(* IEC 61131-3 sources: JingjiangArm/moonboxpro_arm_8.4/Application/Application/数据类型/系统参数/非保持参数, 3 files *)

(* ---- StGrpParam_UnSave.st ---- *)
(*@CES
Name=StGrpParam_UnSave
Type=Gvl
TypeGuid=2db5746d-d284-4425-9f7f-2663a34b0ebc
Guid=502fdab7-460b-44d8-9c01-902a9f3d20a9
HasDeclaration=True
HasImplementation=False
*)
{DECLARATION}
{attribute 'pack_mode' := '1'}
TYPE StGrpParam_UnSave :
STRUCT
	xCutterOnTop_Uw								: BOOL;(* TRUE=放料上裁 *)
	iDebugVelmpm_AxisA_Uw						: INT;(* A轴调试速度/300m/min *)
	iDebugGirthmm_AxisA_Uw						: INT;(* A轴调试周长/300mm *)
	iDebugVelmpm_AxisB_Uw						: INT;(* B轴调试速度/300m/min *)
	iDebugGirthmm_AxisB_Uw						: INT;(* B轴调试周长/300mm *)
	xCutterOnTop_Rw								: BOOL;(* TRUE=收料上裁 *)
	iDebugVelmpm_AxisA_Rw						: INT;(* A轴调试速度/默认300m/min *)
	iDebugGirthmm_AxisA_Rw						: INT;(* A轴调试周长/默认300mm *)
	iDebugVelmpm_AxisB_Rw						: INT;(* B轴调试速度/默认300m/min *)
	iDebugGirthmm_AxisB_Rw						: INT;(* B轴调试周长/默认300mm *)

	xMachineRev									: BOOL;(* 机器反转 *)

	iPromptMsg									: INT;
	iAlarm_TypeId								: INT;//报警轴的类型
	iAlarm_UnitId								: INT;//报警轴位置
	iIdGSE										: INT;
	xFlag_Stop									: BOOL;(* 停机标志/第1次从当前速度降到空转速度，抬所有色组胶辊/牵引速度到0时抬牵引胶辊，第2次按下则将色组从空转停到0速度 *)
	xFlag_PreStart								: BOOL;(* 预启动标志/从停机状态按(预)启动置位标志 色组速度达到空转速度清xFlag_PreStart标志,置位xFlag_Ink标志;当xFlag_Print标志有效后 *)
	xFlag_Ink									: BOOL;(* 匀墨标志/>20m/min不能联动 *)
	xFlag_InkAccing								: BOOL;(* 匀墨加速中<指0~10m/min那个加速过程> *)
	xFlag_Tension								: BOOL;(* 张力投入标志/张力投入有效时收放料变频开始起作用/收放料就位后按印刷按钮,牵引压辊合压/xFlag_Print有效时张力投入不处理 *)
	xFlag_TensionDone							: BOOL;(* 张力ok，可以投入印刷 *)
	xFlag_Print									: BOOL;(* 张力拉料标志有效时，按联动或印刷按钮 先压收牵(延时2s)再压放牵 印刷标志/印刷色组根据联动标志按用户指定的压辊顺序逐一延时压胶辊/胶辊压合完毕后才可置该标志有效 *)
	xFlag_Estop									: BOOL;(* 急停标志/和停机一样要减速到0，只不过减速时间是急停时间 *)
	xFlag_AutoAcc								: BOOL;(* 自动加速 *)
	xFlag_AutoDec								: BOOL;(* 自动减速 *)
	xFlag_ManuAcc								: BOOL;(* 手动加速 *)
	xFlag_ManuDec								: BOOL;(* 手动减速 *)
	xFlag_Accing								: BOOL;(* 加速中 *)
	xFlag_Decing								: BOOL;(* 减速中 *)
	xFlag_EStoping								: BOOL;(* 正在急停中 *)
	xFlag_Stoping								: BOOL;(* 停机中 *)
	xFlag_GotoInking							: BOOL;(* 转到匀墨 *)
	xFlag_InPressing							: BOOL;(* 顺序压辊中 *)
	xFlag_RollerPressDone						: BOOL;(* 压辊处理完成 *)
	xFlag_InchRun								: BOOL;(* 至少有1色处于单运行 *)
	xFlag_AllInchRun							: BOOL;(* 整机单运行标志 *)
	xFlag_AllPress								: BOOL;(* 全体合压 *)
	xFlag_AllUnpress							: BOOL;(* 全体离压 *)
	xFlag_RollerPressAtLeast1					: BOOL;(* 至少1色色组合压 *)
	axFlag_PrnLen_Alarm							: ARRAY [1..3] OF BOOL;(* 计长报警标志 *)
	xFlag_LinkageAxisAlarm						: BOOL;(* 至少有1个联动轴发生报警 *)
	xFlag_TensionUnfinished						: BOOL;(* 张力未完成 *)
	xFlag_VelTooHigh							: BOOL;(* 速度过高 *)
	xFlag_PrestartTimeout						: BOOL;(* 预启动超时标志 *)
	xFlag_KeepAlarming							: BOOL;(* 维持报警*)
	xFlag_ArrivedToTargetVel					: BOOL;(* 到达目标速度 *)
	xFlag_FilmAccDecDone						: BOOL;(* 料膜加减速完成 *)
	xSlowStopTenEn								: BOOL;(* 收放料慢速松料使能/TRUE *)
	xIsDebugMode_Machine						: BOOL;(* 机器调试模式 *)
	uiFilmThickNess								: UINT;(* 料膜厚度/20微米 *)
	abyClrPrnLenCount_Rw						: ARRAY [1..3] OF BYTE;

	iTimeSec_AccDec_AllTheWay					: INT;(* 全程加减速所需要的秒 *)
	rAccDecTime_ThisTime						: REAL;(* 本次加减速时间/单位:s *)

(*2021.11.5.084313/								/ 用于界面显示标准卷径信息 *)
	alrStdVol_Diam_Axis_Hmi						: ARRAY [1..4] OF LREAL;(* 标准卷径值| *)
	alrStdVol_Volt_Axis_Hmi						: ARRAY [1..4] OF LREAL;(* 标准卷径对应的电压值|2019.1.25.142552|更名A轴 *)
	alrStdVol_Coef_Axis_Hmi						: ARRAY [0..4] OF LREAL;(* 分段系数|2019.1.25.142601|更名A轴|[0]表<=1,[1]表>1&& <=2,[2]表>2&& <=3,[3]表>3&& <=4,[4]表>4 *)

	(* 速度 *)
	rVel_Cur									: REAL;(* 当前速度/单位:m/min *)
	rVel_Cur_HMI								: REAL;
	rVel_Film									: REAL;(* 料膜速度/0 *)
	(*											/放料部分 *)
	iSid_AxisA_Uw								: INT;(* 放料站id/-1表示变频/2021.11.21.192354/hdp *)
	xStationOnline_AxisA_Uw						: BOOL;(* 放料a轴驱动器在线标志/2021.12.4.175524/hdp *)
	xMotRev_AxisA_Uw							: BOOL;(* TRUE.放料运动反向/2021.11.21.192354/hdp *)

	iSid_AxisB_Uw								: INT;(* 放料站id/-1表示变频/2021.11.21.192354/hdp *)
	xStationOnline_AxisB_Uw						: BOOL;(* 放料b轴驱动器在线标志/2021.12.4.175524/hdp *)
	xMotRev_AxisB_Uw							: BOOL;(* TRUE.放料运动反向/2021.11.21.192354/hdp *)

	rAI_Uw										: REAL;(* 放料摆臂模拟量输入/-中位值 *)
	rAI_Act_Uw									: REAL;(* 放料摆臂实际模拟量值/2021.11.18.210606 *)
	rAI_HMI_Uw									: REAL;(* 放料摆臂值显示用 *)
	rAI_DiamMeasure_Uw							: REAL;(* 放料卷径测量输入反馈 *)
	arKpid_Current_Uw							: ARRAY [1..3] OF REAL;(* 当前放料pid监控 *)
	stStTimeSet_DnCut_UpCut_Uw_Hmi				: StTimeSet_DnCut_UpCut;(* 放料端的裁切时间集/界面显示 *)
	arKpid_Current_Rw							: ARRAY [1..3] OF REAL;(* 当前收料pid监控 *)
	stStTimeSet_DnCut_UpCut_Rw_Hmi				: StTimeSet_DnCut_UpCut;(* 收料端的裁切时间集/界面显示 *)
	rVel_PreDrv_Uw								: REAL;(* 放料预驱速度 *)
	xReflectionSensorValid_Uw					: BOOL;(* 放料使用弧面信号/FALSE *)
	xReflectSensorLoss_Uw						: BOOL;(* 放料弧面信号丢失标志/FALSE *)
	rDiam_NewVol_Uw								: REAL;(* 放料新卷卷径 *)
	rTowerThetaCur_Uw							: REAL;(* 翻转架当前弧度/0 *)
	rFilmToTowerRollerDis_Uw				: REAL;(*料膜距离导向辊距离|mm*)
	xFilmTouchRoller_Uw						: BOOL;(*料膜接触到了辊子标志*)

	xSts_PreCutting_Uw							: BOOL;(* 放料预备接料/FALSE *)
	rDebugCurVelmpmAxisA_Uw						: REAL;(* A轴调试当前速度/m/min *)
	rDebugCurVelrpmAxisA_Uw						: REAL;(* A轴调试当前速度/r/min *)
	rDebugCurVelmpmAxisB_Uw						: REAL;(* B轴调试当前速度/m/min *)
	rDebugCurVelrpmAxisB_Uw						: REAL;(* B轴调试当前速度/r/min *)

	rDeltaW_RPMIN_Uw							: REAL;(* 放料翻转架转动时候的转速补偿值/0 *)
	xDebugMode_AbsEnc_Uw						: BOOL;(* 放料绝对值编码器调试模式/FALSE *)
	dwAbsEncSinglePos_Uw						: DWORD;(* 放料单圈位置/0 *)
	dwAbsEncSPos_Cur_Uw							: DWORD;(* 放料当前绝对位置/0 *)

	byEncodeValueWr_Uw							: BYTE;(* 放料编码器值写入/放料:01写入轴定位值/02写入A轴最小径定位值/0 *)
	rAIByAbsEnc_Cur_Uw							: REAL;(* 放料绝对值编码器位置转换的电压值/0 *)
	xCutterOnTopFroDebug_Uw						: BOOL;(* 放料上裁刀标志/用于调试/FALSE *)
	xCurAxisAFroDebug_Uw						: BOOL;(* 放料预驱轴为A轴标志/用于调试/FALSE *)
	xAlarmBell_Uw								: BOOL;(* 放料响铃常输出/用于控制定位写入响铃提示使用/FALSE *)
	xIsDebug_DiaMeasure_Uw						: BOOL;(* 放料卷径测量调试模式标志/FALSE *)
	byIsDebug_DiaMeasureArea_Uw					: BYTE;(* 放料卷径测量调试的时候卷径区域值/1 *)
	xIsDebuging_DiaMeasure_Uw					: BOOL;(* 放料卷径测量调试中/FALSE *)
	xCancelDebuging_DiaMeasure_Uw				: BOOL;(* 放料取消卷径测量调试中/FALSE *)
	byAxisDebugBit_Uw							: BYTE;(* 放料轴调试标志/.0\调试使能.1\A轴调试运行.2\A轴自动加减速.3\A轴运行中.4\B轴调试运行.5\B轴自动加减速.6\B轴运行中/0 *)
	byAxisDebugBit_Uw_2							: BYTE;(* 放料2轴调试标志/.0\调试使能.1\A轴调试运行.2\A轴自动加减速.3\A轴运行中.4\B轴调试运行.5\B轴自动加减速.6\B轴运行中/0 *)
	xEnCodeErr_Uw								: BOOL;(* 放料编码器故障*)
	xEnCodeErr_Rw								: BOOL;(* 收料编码器故障*)

	rPi_Value_Uw								: REAL;(* 放料pi值/0 *)
	rForwardStep_Uw								: REAL;(* 放料升降速前馈/0 *)
	rTotalPiValue_Uw							: REAL;
	xAxisAForeward_Uw							: BOOL;(* 放料A轴正转/FALSE *)
	xAxisBForeward_Uw							: BOOL;(* 放料B轴正转/FALSE *)
	rVelRPM_Cur_Uw								: REAL;(* 放料当前转速/0 *)
	rAxisAVelRPM_Cur_Uw							: REAL;(* 放料A轴转速/0/2021.11.18.201209 *)
	rAxisBVelRPM_Cur_Uw							: REAL;(* 放料B轴转速/0/2021.11.18.201209 *)
	xFlag_DiamCalc_ing_Uw						: BOOL;(* 放料卷径计算中 *)
	xFlag_DiamCalc_end_Uw						: BOOL;(* 放料卷径计算完成 *)
	xFlag_DiamMeasure_end_Uw					: BOOL;(* 放料卷径测量完成 *)
	xFlag_PreDrv_ing_Uw							: BOOL;(* 放料预驱中... *)
	xFlag_PreDrv_end_Uw							: BOOL;(* 放料预驱完成  *)
	xFlag_Cut_ing_Uw							: BOOL;
	xFlag_Cut_end_Uw							: BOOL;
	xFlag_VolDiamAlarm_Uw						: BOOL;(* 卷径报警标志 *)
	rAI_DiamMeasure_HMI_Uw						: REAL;(* 兼容摆臂输入类型转换后的卷径测量结果屏显值/2021.11.5.175329 *)
	xAITypeBtn_Uw								: BOOL;(* 输入类型切换按钮/2021.11.18.201254 *)

	(*											/收料部分 *)
	iSid_AxisA_Rw								: INT;(* 收料站id/-1表示变频/2021.11.21.192354/hdp *)
	xStationOnline_AxisA_Rw						: BOOL;(* 收料a轴驱动器在线标志/2021.12.4.175524/hdp *)
	xMotRev_AxisA_Rw							: BOOL;(* TRUE.收料运动反向/2021.11.21.192354/hdp *)

	iSid_AxisB_Rw								: INT;(* 收料站id/-1表示变频/2021.11.21.192354/hdp *)
	xStationOnline_AxisB_Rw						: BOOL;(* 收料b轴驱动器在线标志/2021.12.4.175524/hdp *)
	xMotRev_AxisB_Rw							: BOOL;(* TRUE.收料运动反向/2021.11.21.192354/hdp *)

	rAI_Rw										: REAL;(* 收料摆臂模拟量输入/-中位值 *)
	rAI_Act_Rw									: REAL;(* 收料摆臂实际模拟量值/2021.11.18.201450 *)
	rAI_HMI_Rw									: REAL;(* 收料摆臂值显示用 *)
	rVel_PreDrv_Rw								: REAL;(* 收料预驱速度 *)
	rDiam_NewVol_Rw								: REAL;(* 收料新卷卷径 *)
	rTaper_Rw									: REAL;(* 收料锥度 *)

	xSts_PreCutting_Rw							: BOOL;(* 收料预备接料 *)
	rDebugCurVelmpmAxisA_Rw						: REAL;(* A轴调试当前速度/m/min *)
	rDebugCurVelrpmAxisA_Rw						: REAL;(* A轴调试当前速度/r/min *)

	rDebugCurVelmpmAxisB_Rw						: REAL;(* B轴调试当前速度/m/min *)
	rDebugCurVelrpmAxisB_Rw						: REAL;(* B轴调试当前速度/r/min *)
	xDebugMode_AbsEnc_Rw						: BOOL;(* 收料绝对值编码器调试模式/默认FALSE *)
	dwAbsEncSinglePos_Rw						: DWORD;(* 收料单圈位置/0 *)
	dwAbsEncSPos_Cur_Rw							: DWORD;(* 收料当前绝对位置/0 *)
	byEncodeValueWr_Rw							: BYTE;(* 收料编码器值写入/收料/01写入轴定位值/0 *)
	xCutterOnTopFroDebug_Rw						: BOOL;(* 收料上裁刀标志/用于调试/FALSE *)
	xCurAxisAFroDebug_Rw						: BOOL;(* 收料预驱轴为A轴标志/用于调试/FALSE *)
	x6InchFroDebug_Rw       					: BOOL;(* 收料6寸标志/用于调试/FALSE*)
	xAlarmBell_Rw								: BOOL;(* 收料响铃常输出/用于控制定位写入响铃提示使用/FALSE *)
	byAxisDebugBit_Rw							: BYTE;(* 收料轴调试标志/.0\调试使能.1\A轴调试运行.2\A轴自动加减速.3\A轴运行中.4\B轴调试运行.5\B轴自动加减速.6\B轴运行中/0 *)
	rPi_Value_Rw								: REAL;(* 收料pi值/0 *)
	rForwardStep_Rw								: REAL;(* 收料升降速前馈/0 *)
	rTotalPiValue_Rw							: REAL;
	xAxisAForeward_Rw							: BOOL;(* 收料A轴正转/FALSE *)
	xAxisBForeward_Rw							: BOOL;(* 收料B轴正转/FALSE *)
	rVelRPM_Cur_Rw								: REAL;(* 收料当前转速/0 *)
	rAxisAVelRPM_Cur_Rw							: REAL;(* 收料A轴转速/0/2021.11.18.201604 *)
	rAxisBVelRPM_Cur_Rw							: REAL;(* 收料B轴转速/0/2021.11.18.201608 *)
	xFlag_6Inch_Rw								: BOOL;(* 收料6寸标志/反之为3寸/FALSE *)
	xFlag_PreDrv_ing_Rw							: BOOL;(* 收料预驱中... *)
	xFlag_PreDrv_end_Rw							: BOOL;(* 收料预驱完成 *)
	xFlag_Cut_ing_Rw							: BOOL;(* 收料裁切中 *)
	xFlag_Cut_end_Rw							: BOOL;(* 收料裁切完成 *)
	xAITypeBtn_Rw								: BOOL;(* 输入类型切换按钮 *)

	(*											/放牵部分 *)
	iSid_If										: INT;(* 放牵站id/-1表示变频 *)
	xStationOnline_If							: BOOL;(* 放牵驱动器在线标志/2021.12.4.175524/hdp *)
	xMotRev_If									: BOOL;(* TRUE.放牵运动反向/2021.11.16.134652/+ *)
(* 2021.12.29.153030/hdp *)

	rAI_If										: REAL;(* 放牵摆臂模拟量输入/-中位值 *)
	rAI_Act_If									: REAL;(* 放牵摆臂实际模拟量值/2021.11.18.201802 *)
	rAI_HMI_If									: REAL;(* 放牵摆臂值显示用 *)
	xInchBtn_If									: BOOL;(* 放牵单运行/FALSE *)
	xRollerSts_If								: BOOL;(* 放牵压辊/FALSE *)
	xRunEn_If									: BOOL;(* 放牵运动使能/0/2021.11.18.201925 *)
	rVel_Cur_If									: REAL;(* 放牵速度/0 *)
	rPi_Value_If								: REAL;(* 放牵pi值/0 *)
	rForwardStep_If								: REAL;(* 放牵升降速前馈/0 *)
	rUsingGirth_If								: REAL;(* 放牵速度控制实际使用的周长/500mm *)
	xInching_If									: BOOL;(* 放牵单运行中/FALSE *)
	xAITypeBtn_if								: BOOL;(* 输入类型切换按钮 *)
	(*											/收牵部分 *)
	iSid_Of										: INT;(* 收牵站id/-1表示变频 *)
	xStationOnline_Of							: BOOL;(* 收牵驱动器在线标志/2021.12.4.175524/hdp *)
	xMotRev_Of									: BOOL;(* TRUE.收牵运动反向/2021.11.16.134652/+ *)

	rAI_Of										: REAL;(* 收牵摆臂模拟量输入/-中位值 *)
	rAI_Act_Of									: REAL;(* 收牵摆臂实际模拟量值/2021.11.18.202051 *)
	rAI_HMI_Of									: REAL;(* 收牵摆臂值显示用 *)
	xInchBtn_Of									: BOOL;(* 收牵单运行/FALSE *)
	xRollerSts_Of								: BOOL;(* 收牵压辊/FALSE *)
	xRunEn_Of									: BOOL;(* 收牵运动使能/0/2021.11.18.202215 *)
	rVel_Cur_Of									: REAL;(* 收牵速度/0 *)
	rPi_Value_Of								: REAL;(* 收牵pi值/0 *)
	rForwardStep_Of								: REAL;(* 收牵升降速前馈/0 *)
	rUsingGirth_Of								: REAL;(* 收牵速度控制实际使用的周长/500mm *)
	xInching_Of									: BOOL;(* 收牵单运行中/FALSE *)
	xAITypeBtn_Of								: BOOL;(* 输入类型切换按钮/2021.11.18.202322 *)
	sCurRecipeName_InUse							: STRING ;(*当前加在的配方*)
	dwSTS_ALL									: DWORD;(* 2021.11.4.174929 *)
(*												/ 整机状态 *)
(*												/bit0.整机套印纵向自动 *)
(*												/bit1.整机套印横向自动 *)
(*												/*)
(*												/bit8.主站的通讯记录到日志中 *)
(*												/*)
(*												/*)
(*												/bit16.主站请置该标志有效/2021.11.6.102700 *)
(*												/bit17.置位标识显示精采样波形 *)
(*												/*)
(*												/*)
(*												/*)
(*												/bit24.dll显示调试信息/2021.12.1.191835/hdp *)
(*												/bit25.精采样显示阀值3 *)
(*												/bit26.精采样显示阀值2 *)
(*												/bit27.精采样显示阀值1 *)
(*												/bit28.精采样显示峰值位置 *)
(*												/bit29.精采样显示最小值位置 *)
(*												/bit30.精采样显示最大值位置 *)
(*												/bit31.精采样显示基线 *)

	xAutoAccDec_Hmi								: BOOL;
	xFlag_IfOf_Ink								: BOOL;(*空转牵引联动标志*)
	xFlag_FastStoping						: BOOL;
	rFinalVelocity							: REAL;(*末速度*)

	xFlag_AutoMaticCutting_Uw					: BOOL;(*2022.4.25.090246 自动裁切中标志*)
(*	abyReserved1							: ARRAY [1..4] OF BYTE;*)
	xFlag_AutoMaticCutting_rw					: BOOL;(*2022.4.25.090246 自动裁切中标志*)
	rAutoMaticCuttingLenth_CurMode_uw			: REAL;(*放料自动裁切当前模式下的计米值|2022.4.26.101850*)
	rActRemainFilmLenth_Uw						: REAL;(*实际剩余长度|mm-测量值*)
	rAutoMaticCuttingLenth_CurMode_Rw			: REAL;(*收料自动裁切当前模式下的计米值|2022.4.26.101850*)

	xCurAxisDia_Uw_Wr							: BOOL;(*写入当前轴的卷径|2022.4.9.230449*)
	xCurAxisDia_Rw_Wr							: BOOL;(*写入当前轴的卷径|2022.4.9.230449*)
	rTaper_Cur_Uw								: REAL;(*锥度当前|放料|*)
	rTaper_Cur_If								: REAL;(*锥度当前|放牵|*)
	rTaper_Cur_Of								: REAL;(*锥度当前|收牵|*)

	rTaperValueBegin_Hmi_Uw						: REAL;(*放料起始锥度显示值|根据单位切换*)
	rTaperValueEnd_Hmi_Uw						: REAL;(*放料结束锥度显示值|根据单位切换*)
	rTaperValueBegin_Hmi_Rw						: REAL;(*收料起始锥度显示值|根据单位切换*)
	rTaperValueEnd_Hmi_Rw						: REAL;(*收料结束锥度显示值|根据单位切换*)
	rTaperValueBegin_Hmi_If						: REAL;(*放牵起始锥度显示值|根据单位切换*)
	rTaperValueEnd_Hmi_If						: REAL;(*放牵结束锥度显示值|根据单位切换*)
	rTaperValueBegin_Hmi_Of						: REAL;(*收牵起始锥度显示值|根据单位切换*)
	rTaperValueEnd_Hmi_Of						: REAL;(*收牵结束锥度显示值|根据单位切换*)

	byTaperUnitConfirm_Uw						: BYTE;(*放料锥度单位确认|.0 N确认|.1 Mpa确认*)
	byTaperUnitConfirm_Rw						: BYTE;(*收料锥度单位确认|.0 N确认|.1 Mpa确认*)
	byTaperUnitConfirm_If						: BYTE;(*放牵锥度单位确认|.0 N确认|.1 Mpa确认*)
	byTaperUnitConfirm_Of						: BYTE;(*收牵锥度单位确认|.0 N确认|.1 Mpa确认*)
	(*2021.7.29.105859 增加|16BYTES*)
	rTaperValueCur_Hmi_If						: REAL;(*放牵锥度当前值|根据单位切换*)
	rTaperValueCur_Hmi_of						: REAL;(*收牵锥度当前值|根据单位切换*)
	rTaperValueCur_Hmi_Uw						: REAL;(*放料锥度当前值|根据单位切换*)
	rTaperValueCur_Hmi_Rw						: REAL;(*收料锥度当前值|根据单位切换*)
	rValue_DiaMeasure							: REAL;(*卷径测量采样值*)
	rVolt_CalcDiam_Used_Watch					: REAL;(*计算卷径的电压值*)
	rAO_Inverter_Uw_AxisA						: REAL;(*放料A轴输出|2017-08-12 17:25:33*)
	rAO_Inverter_Uw_AxisB						: REAL;(*放料B轴输出|2017-08-12 17:25:33*)
	rAO_Inverter_Rw_AxisA						: REAL;(*收料A轴输出|2017-08-12 17:25:33*)
	rAO_Inverter_Rw_AxisB						: REAL;(*收料B轴输出|2017-08-12 17:25:33*)

	xBtn_HorzPreRegister_Repeat				: BOOL;(*横向重复值按钮*)
	xBtn_HorzPreRegister_Setup				: BOOL;(*横向设定值按钮*)
	xSts_HorzPreRegister					: BOOL;(*横向预套准状态*)
	xMode_HorzPreRegister					: BOOL;(*横向预套准方式：FALSE为设定值;TRUE是重复值*)
	xFlag_HorzPreRegister_All_end			: BOOL;(*横向预套准全部完成*)
	xFlag_Home								: BOOL;
	xFlag_Home_ing							: BOOL;
	xFlag_Home_end							: BOOL;
	xFlag_ConfirmPreRegHomePos				: BOOL;(*2017-09-13 12:51:52| 确认预套准基准点*)
	xFlag_ConfirmPreRegHomePos_ing			: BOOL;(*确认预套准基准点-ing*)
	xFlag_ConfirmPreRegHomePos_end			: BOOL;(*确认预套准基准点-end*)
	xFlag_PreRegister						: BOOL;
	xFlag_PreRegister_ing					: BOOL;
	xFlag_PreRegister_end					: BOOL;
	xFlag_PhaseRestore						: BOOL;(*相位恢复*)
	xFlag_PhaseRestore_ing					: BOOL;(*相位恢复-ing*)
	xFlag_PhaseRestore_end					: BOOL;(*相位恢复-end*)
	xBtn_Home								: BOOL;
	xBtn_ConfirmPreRegHomePos				: BOOL;
	xBtn_PreRegister						: BOOL;
	xBtn_PhaseSave							: BOOL;(*相位保存*)
	xBtn_PhaseRestore						: BOOL;(*相位恢复*)
	xFlag_MotionParamInitialized				: BOOL;(*加速度初始化完成-计算加速度目标速度加加速度*)
	xFlag_AccDecStop							: BOOL;
	//下面时牵引收放料中心辊的离线报警位置偏差报警标志
	xNetOffline_CENTRAL:BOOL;
	xAxisAlarm_CENTRAL:BOOL;
	xPosDeviationAlarm_CENTRAL:BOOL;
	xNetOffline_CENTRAL2:BOOL;
	xAxisAlarm_CENTRAL2:BOOL;
	xPosDeviationAlarm_CENTRAL2:BOOL;
	xNetOffline_IF:BOOL;
	xAxisAlarm_IF:BOOL;
	xPosDeviationAlarm_IF:BOOL;
	xNetOffline_OF:BOOL;
	xAxisAlarm_OF:BOOL;
	xPosDeviationAlarm_OF:BOOL;
	xNetOffline_UW_A:BOOL;
	xAxisAlarm_UW_A:BOOL;
	xPosDeviationAlarm_UW_A:BOOL;
	xNetOffline_UW_B:BOOL;
	xAxisAlarm_UW_B:BOOL;
	xPosDeviationAlarm_UW_B:BOOL;
	xNetOffline_RW_A:BOOL;
	xAxisAlarm_RW_A:BOOL;
	xPosDeviationAlarm_RW_A:BOOL;
	xNetOffline_RW_B:BOOL;
	xAxisAlarm_RW_B:BOOL;
	xPosDeviationAlarm_RW_B:BOOL;
	//2023.8.18.143718具体报警信息
	dwAlarmDetail_CENTRAL:DWORD;//轴报警信息-ZHONGX
	dwAlarmDetail_CENTRAL2:DWORD;//轴报警信息-ZHONGX

	dwAlarmDetail_IF:DWORD;//轴报警信息-放牵
	dwAlarmDetail_OF:DWORD;//轴报警信息-收前
	dwAlarmDetail_UW_A:DWORD;//轴报警信息-放A
	dwAlarmDetail_UW_B:DWORD;//轴报警信息-放B
	dwAlarmDetail_RW_A:DWORD;//轴报警信息-收A
	dwAlarmDetail_RW_B:DWORD;//轴报警信息-收B

	xValid_CentralDrum							: BOOL;(* 中心滚筒有效标志 *)
	iSid_CentralDrum							: INT;(* 中心滚筒站id/初始-1/有效性通过查表确定 *)
	xStationOnline_CentralDrum					: BOOL;(* 站在线标志-中心滚筒/读取站号以后实时更新 *)
	xMotRev_CentralDrum							: BOOL;(* 中心滚筒电机反向运动 *)
	rAxisVel_CentralDrum						: REAL;(* 中心滚筒轴速度 *)
	xPrintInching: BOOL;//整机点动
	rVel_Inching_Print: REAL;//点动速度
	xTapPosition_Breaking					: BOOL;(*断料档位|*)
	xTapPosition_UniformInk					: BOOL;(*匀墨档位|*)
	xTapPosition_Printing					: BOOL;(*印刷档位|*)
	wEn_UwRw_IfOf_Center					: WORD;(*牵引收放料中心辊的使能标志*)
											(*bit0:放牵*)
											(*bit1:收牵*)
											(*bit2:放A*)
											(*bit3:放B*)
											(*bit4:收A*)
											(*bit5:收B*)
											(*bit6:中心辊1*)
											(*bit7:中心辊2*)
	aiMotionStep_AllStation					: ARRAY [1..MAX_STATION_NUM] OF INT;
	byBtn_ConfirmMedian						: BYTE;
	xUwVolDiamMeasurementFailed								: BIT;(*放料卷径检测失败*)
	xBtnClrAlarmInf											: BIT;(*报警清楚按钮*)

	byPseudoRandomId						: BYTE:=1;(*=0 放牵|=1 放料|=2 收料 |=3 收牵*)
	xPseudoRandomEn							: BOOL;(*伪随机使能*)
	aiTestPseudoRandom_Kp					: ARRAY [1..3] OF INT;(*伪随机测试Kp*)
	aiTestPseudoRandom_Kd					: ARRAY [1..3] OF INT;(*伪随机测试Kd*)
	xPseudoRandomTsting						: BOOL;(*伪随机测试中*)
	xDebug_Enc_Uw							: BOOL;(*放料调试*)
	xDebug_Enc_Rw							: BOOL;(*收料调试*)
	wAxisDebug_UwRw							: WORD;(*轴调试标志|.0\放料调试使能.1\放料A轴调试运行.2\放料A轴自动加减速.3\放料A轴运行中.4\放料B轴调试运行.5\放料B轴自动加减速.6\放料B轴运行中
									  .8\收料调试使能.9\收料A轴调试运行.10\收料A轴自动加减速.11\收料A轴运行中.12\收料B轴调试运行.13\收料B轴自动加减速.14\收料B轴运行中*)
	xFlag_SafeTyGratingProctec_Uw			: BOOL;(*放料光栅保护标志*)
	xFlag_SafeTyGratingProctec_Rw			: BOOL;(*放料光栅保护标志*)

	bySetTestPid_IfOf:BYTE;(*设置伪随机测试的pid值*)
	bySetTestPid_Uw:BYTE;(*设置伪随机测试的pid值*)
	bySetTestPid_Rw:BYTE;(*设置伪随机测试的pid值*)
	bySetTestPid_If:BYTE;(*设置伪随机测试的pid值*)
	bySetTestPid_Of:BYTE;(*设置伪随机测试的pid值*)
	xLinkage_IfOf_Ink: BOOL;
	xFlag_Cut_end_Uw_UseInOtherPrg: BOOL;
	xFlag_Cut_ing_Uw_UseInOtherPrg: BOOL;
	xFlag_Cut_end_Rw_UseInOtherPrg: BOOL;
	xConfirmRad0: BOOL;(*0弧度确认*)
	xFlag_Follow_1U_V_UwCut		: BOOL;(*裁切跟一色标志*)
	xKeepAlarm_NoMaterial			: BOOL;(*没料持续报警*)
	xKnob_6Inch_Rw				: BOOL;(*界面收料6吋切换开关*)
	xWillAutoMaticPreCut_Uw		: BOOL;(**)
	axMeasure_StdVol						: ARRAY [1..4] OF BOOL;(*卷径测量按钮*)
	rPseudoRandomRoundAmplitude_Cur		: REAL;

	rAxisAFreq_Uw						: REAL;(*放料A频率监控*)
	rAxisBFreq_Uw						: REAL;(*放料A频率监控*)
	rAxisAFreq_Rw						: REAL;(*放料A频率监控*)
	rAxisBFreq_Rw						: REAL;(*放料A频率监控*)

	xAllowSwitchCutter_Uw				: BOOL;(*收放料允许切换上下裁刀标志@|./0 放料可以|./1 收料可以*)
	xAllowSwitchCutter_Rw				: BOOL;(*收放料允许切换上下裁刀标志@|./0 放料可以|./1 收料可以*)
	xAxisALocation_Use_Uw					: BOOL;
	xAxisBLocation_Use_Uw					: BOOL;
	xAxisALocation_Use_Rw					: BOOL;
	xAxisBLocation_Use_Rw					: BOOL;

	rWuCompensate_Uw:REAL;(*补偿的转速(R/MIN)|计算的*)
	rWuCompensate_Act_Uw:REAL;(*补偿的转速(R/MIN)|实际使用的*)

	rWuCompensate_Rw:REAL;(*补偿的转速(R/MIN)|计算的*)
	rWuCompensate_Act_Rw:REAL;(*补偿的转速(R/MIN)|实际使用的*)
	rTaperMax_Uw: REAL;
	rTaperMax_Rw: REAL;
	rTaperMax_If: REAL;
	rTaperMax_Of: REAL;

	xGirthCalFinish_If: BOOL;
	xGirthCalFinish_Of: BOOL;
	(*扰动输出的控制输入参数@2024.12.3.102359*)
	xEn_Disturbance_If: BOOL;(*扰动使能*)
	rFreq_Disturbance_If: REAL:=1;(*扰动频率@hz*)
	rAmplitude_Disturbance_If:REAL:=1;(*扰动幅值*)
	uiTotalTime_Disturbance_If: UINT:=0;(*扰动输出的总时间|=0 代表一直输出@s*)
	xOuting_sin_If:BOOL:=FALSE;(*输出标志*)
	rResult_sin_If: REAL:=0;
	xEn_Disturbance_Of: BOOL;(*扰动使能*)
	rFreq_Disturbance_Of: REAL:=1;(*扰动频率@hz*)
	rAmplitude_Disturbance_Of:REAL:=1;(*扰动幅值*)
	uiTotalTime_Disturbance_Of: UINT:=0;(*扰动输出的总时间|=0 代表一直输出@s*)
	xOuting_sin_Of:BOOL:=FALSE;(*输出标志*)
	rResult_sin_Of: REAL:=0;
	rVelRPM_Cur_If: REAL;(*放牵转速*)
	rVelRPM_Cur_Of: REAL;(*收牵转速*)
	byPseudoRandomRoundTimes_Cur: BYTE;(*伪随机测试当前次数*)
	xFlagFollow1U_AccDecing: BOOL;(*加减速跟踪第一色标志*)
	byGrpArcAxisNum			: BYTE;
	abyGrpArcAxisList: ARRAY [1..MAX_UNIT_NUM] OF BYTE;
	abyGrpFollowArcIdList: ARRAY [1..MAX_UNIT_NUM] OF BYTE;
	abyGrpArcIdList	: ARRAY [1..MAX_UNIT_NUM] OF INT;
	xEnaTestARC_Ink							: BOOL;(*空转测试使能*)
	rAcceleration_Max				: REAL;(*最大加速度*)
	rAcceleration_Cur				: REAL;(*当前加速度*)

	byGrpAxisNum_Pu					: BYTE;
	abyGrpAxisList					: ARRAY [1..MAX_UNIT_NUM] OF BYTE;
	iAxisId_StepTest_V						: INT;(*阶跃测试的轴id*)
	iMicron_StepTest1_V						: INT;(*阶跃测试的数值|单位:um*)
	iMicron_StepTest2_V						: INT;(*阶跃测试的数值|单位:um*)
	iInterval_StepTest12					: INT;(*2此阶跃的间隔|幅*)

	xSwitch_AutoAdjust_V_Grp				: BIT;(*整机手自动*)
	xSwitch_AutoAdjust_H_Grp				: BIT;(*整机手自动*)
	xLinkage_If								: BIT;(*放牵联动*)
	xLinkage_Of								: BIT;(*收牵联动*)
	xMoveEnable_Motor_If					: BIT;
	xMoveEnable_Motor_Of					: BIT;
	rMainVel_Uw : REAL;
	rMainVel_Rw : REAL;

	(*2025.8.13.103441||新增工艺参数*)
	lrAxisScraperVel:LREAL;
	rHz_UnitScraper_CurrWR: REAL;(*刮刀速度写入变频值-485变频*)
	rHz_UnitInkRoller_CurrWR: REAL;

	(*2025.08.13.145324 || 至少联动一色标志*)
	xFlag_LinkageAtleast1Axis					: BOOL;
	(*新增变量-开始|wang.nt|2025.08.13.144038*)
	xWillAutoMaticPreCut_Rw : BOOL;(*收料即将自动接料*)
	xFlag_HotBlowerStopDelay : BOOL;(*热风延时关闭中*)
	xInverterAlarmCurAxis_Uw				: BOOL;(*放料变频器当前轴报警*)
	xInverterAlarmCurAxis_Rw				: BOOL;(*收料变频器当前轴报警*)
	xInverterAlarmPreAxis_Uw				: BOOL;(*放料变频器预驱轴报警*)
	xInverterAlarmPreAxis_Rw				: BOOL;(*收料变频器预驱轴报警*)
	xFlag_FastStopBtnDn:BOOL;(*快停被按下|2022.4.13.155130*)
	xEstopBtnDne:BOOL;(*急停被按下*)
	xTowerInvAlarm_Uw:BOOL;
	xTowerInvAlarm_Rw:BOOL;
	xInverterAlarm_If				: BOOL;(*放牵变频器报警*)
	xInverterAlarm_Of				: BOOL;(*收牵变频器报警*)
	(*新增变量-结束|wang.nt|2025.08.13.144054*)

	xBtn_StepTest_V							: BOOL;(*纵向阶跃*)

(*2025.8.20.200913*)
	xBtn_ExhAir_Reset						: BIT;(*排风复位按钮*)
	xBtn_CopyExhFreq_1U_To_Other			: BIT;(*复制1U排风频率到所有色*)
	xBtn_AllExhAir_Off						: BIT;(*全体排风关*)
	xBtn_AllExhAir_On						: BIT;(*全体排风开*)
	xBtn_Reset_TempCtlBlock					: BIT;(*复位温控模块按钮*)
	xBtn_CopySV_1U_To_Other					: BIT;(*复制1U排风频率到所有色*)
	xBtn_AllHeating_Elc						: BIT;(*全体电加热*)
	xBtn_AllHeating_I						: BIT;(*全体加热I当*)
	xBtn_AllHeating_II		  				: BIT;(*全体加热II当*)
	xBtn_AllHeating_III					    : BIT;(*全体加热III当*)
	xBtn_AllHeating_Close					: BIT;(*全体加热关*)
	xBtn_AllHeating_Water	 			    : BIT;	(*全体水加热*)
	(*预套准相关变量|wang.nt|2025.08.21.171436*)
	xFlag_PhaseSave:BOOL;(*固定相位保存相关|2024.9.6.213011*)
	xFlag_PhaseSave_end:BOOL;
	xFlag_PhaseRead:BOOL;
	xFlag_PhaseRead_end:BOOL;
	xBtn_SaveAllData:BOOL;(*全部参数保存|不管有没有都写入一次当前值*)
	xBtn_SaveProtionData:BOOL;(*部分参数保存|没有相位值的色组*)
	xBtn_SaveCancel:BOOL;(*界面关闭*)
	xFlag_AxisInitPhaseHmiDis:BOOL;(*轴的初始相位操作界面显示*)
	byFirstValidAxisId						: BYTE;(*2018.9.9.203836\首个有效轴|*)

	(*2025.9.25.110708从这开始是润新测试完后增加内容*)
	iStationId_Alarm: INT;(*报警时给这个变量赋值-无报警时赋值255吧*)
	abyAxisList_CoatingPrn					: ARRAY [1..MAX_UNIT_NUM] OF BYTE;(*涂布轴列表|*)
	byAxisNum_CoatingPrn					: BYTE;
	xInching_Uw: BOOL;
	xInching_Rw: BOOL;
	xArcErrInRange: BOOL;
	rAIMax_Uw: REAL;
	rAIMin_Uw: REAL;
	rAIMax_Rw: REAL;
	rAIMin_Rw: REAL;
	rAIMin_If: REAL;
	rAIMax_If: REAL;
	rAIMin_Of: REAL;
	rAIMax_Of: REAL;

(*2025.11.5.154018*)
	xBtn_PreRegisterAxisId_Manu					: BIT;(*预套准的轴号手动确定@不考虑联动开关*)
	xBtn_PreRegisterCorrConfirm: BIT;//预套准自动修正按钮

	//xRsv_Flag4										: BIT;
	//xRsv_Flag5										: BIT;
	//xRsv_Flag6										: BIT;
	//xRsv_Flag7										: BIT;
	//再取一个BYTE用做BIT||4-1=3
	//2025.10.20.153729||bit0和bit1用作横向预套准按钮
//2025.12.31.111752增加变量，数据结构变化
	rCur_PressureValue	: REAL;//牵引压力传感器当前值

END_STRUCT
END_TYPE

{IMPLEMENTATION}

(* ---- StSysParam_UnSave.st ---- *)
(*@CES
Name=StSysParam_UnSave
Type=Gvl
TypeGuid=2db5746d-d284-4425-9f7f-2663a34b0ebc
Guid=a407ba0f-c9c2-422c-ab5e-e61307b67d21
HasDeclaration=True
HasImplementation=False
*)
{DECLARATION}
{attribute 'pack_mode' := '1'}
TYPE StSysParam_UnSave :
STRUCT
	stStSysCfgStruct							: StSysCfgStruct;(* 2022.6.8.154438/hdp/系统配置更改结构 *)
	byCurrUsrLevel								: BYTE;(*用户等级处理*)
	diEncPos_Virtual							: DINT;
	(*tcp需要的*)
	(*[2]=厂家支持设备@10bytes*)
	xCommEn_Tcp:BOOL;(*厂家支持设备tcp通讯使能@常有效*)
	xOpenSocketing:BOOL;(*厂家支持设备tcp打开中@连接中*)
	xOpenSocketDne:BOOL;(*厂家支持设备tcp打开成功*)
	xOpenSocketFailed:BOOL;(*厂家支持设备tcp打开失败*)
	xConnectOk_Tcp: BOOL;(*厂家支持设备连接成功了*)
	byConnectSts_Tcp:BYTE;(*厂家支持设备的连接状态		  @=0 未打开
														  @=1 打开中@连接中
														  @=2 打开成功
														  @=3 打开失败
														  @=4 通讯超时*)
	abyReserved_Tcp:ARRAY [1..4] OF BYTE;

	(*[1]=监控设备@10bytes*)
	xCommEn_WatchDevice_Tcp:BOOL;(*监控设备tcp通讯使能@常有效*)
	xOpenSocketing_WatchDevice:BOOL;(*监控设备tcp打开中@连接中*)
	xOpenSocketDne_WatchDevice:BOOL;(*监控设备tcp打开成功*)
	xOpenSocketFailed_WatchDevice:BOOL;(*监控设备tcp打开失败*)
	xConnectOk_WatchDevice_Tcp: BOOL;(*监控设备连接成功了*)
	byConnectSts_WatchDevice_Tcp:BYTE;(*监控设备的连接状态@=0 未打开
														  @=1 打开中@连接中
														  @=2 打开成功
														  @=3 打开失败
														  @=4 通讯超时*)
	abyReserved1_Tcp:ARRAY [1..4] OF BYTE;

(*新增2023.10.14.104239||11字节*)
	(*485需要的@10bytes*)
	xCommEn_485:BOOL;(*485通讯使能开关*)
	xOpenPortDne:BOOL;(*485打开成功*)
	xOpenPortFailed:BOOL;(*485打开失败*)
	xCommEn_WatchDevice_485:BOOL;(*监控设备通讯使能*)
	byConnectSts_485:BYTE;(*485设备的连接状态@=0 未打开
											 @=1 打开中@连接中@485不用
											 @=2 打开成功
											 @=3 打开失败*)
	abyReserved_485:ARRAY [1..5] OF BYTE;

	rAO0_WaterValue_Start					: REAL;
	rAO0_WaterValue_Start2					: REAL;

	dwCtl_FromDiamonds						: DWORD;(*金刚界面的一些临时按钮控制*)
											(*
											bit0~bit15: A系用
											bit0: 预启动
											bit1: 停机
											bit2: 急停
											bit16~bit31: B系用
											bit16: 预启动
											bit17: 停机
											bit18: 急停
											*)
	byTaperUnitType:BYTE;(*张力单位切换标志|.0 放牵\.1收牵\.2放料\.3收料*)
	byCurGrpId_HMI: BYTE;(*当前界面的系号*)
	byArcDeCoupleStepTest:BYTE;(*套色阶跃测试@=1 经过小黄解耦控制器输出阶跃调整量
											   @=2 不经过解耦控制器直接阶跃输出*)
	xSaveFineSampleData_ToArc: BOOL;
	iAxisId_CurSmpData: INT;(*当前显示的波形机组号*)
	abyData_T1_R: ARRAY [1..4000] OF BYTE;
	abyData_T1_G: ARRAY [1..4000] OF BYTE;
	abyData_T1_B: ARRAY [1..4000] OF BYTE;
	abyData_T2_R: ARRAY [1..4000] OF BYTE;
	abyData_T2_G: ARRAY [1..4000] OF BYTE;
	abyData_T2_B: ARRAY [1..4000] OF BYTE;

	aiStationList_UnitController: ARRAY [1..MAX_STATION_NUM] OF INT;(*用月光宝盒/PRO时候，需要一个控制器列表，用于通讯？*)
	aiAxisIdList_UnitArcAdj: ARRAY [1..MAX_STATION_NUM] OF INT;(*用月光宝盒/PRO时候，需要一个轴列表-对应宝盒/PRO*)

	(*2025.8.19.213305*)
	dwAxis_SkipTheHeader				: DWORD;(*让料头标志| 位标志bit0=机组1,...,bit31=机组32*)

	xIOTestMode: BIT;(*IO测试模式*)
	xMoveFreq_I_ToAll_AirHot: BIT;
	xMoveFreq_II_ToAll_AirHot: BIT;
	xMoveFreq_III_ToAll_AirHot: BIT;
	xMoveFreq_I_ToAll_ExhaustAir: BIT;
	xMoveFreq_II_ToAll_ExhaustAir: BIT;
	xMoveFreq_III_ToAll_ExhaustAir: BIT;
	xSwitch_ScraperReset								: BIT;
	xSwitch_InkRollerReset								: BIT;
	xSwitch_HotwindReset: BIT;
	xSwitch_ResetTemctlModule: BIT;
	xSwitch_Copy1stUExhaustDamperPos : BIT;
	xInkGrooveCali_Hmi: BIT;

END_STRUCT
END_TYPE

{IMPLEMENTATION}

(* ---- StUnitParam_UnSave.st ---- *)
(*@CES
Name=StUnitParam_UnSave
Type=Gvl
TypeGuid=2db5746d-d284-4425-9f7f-2663a34b0ebc
Guid=be979c59-c798-41af-9e86-c1d3d1a3e0f0
HasDeclaration=True
HasImplementation=False
*)
{DECLARATION}
{attribute 'pack_mode' := '1'}
TYPE StUnitParam_UnSave :
STRUCT
	xMotRev_BottomRoller						: BOOL;(* 底辊电机反向运动 *)
	xSamRev_BottomRoller						: BOOL;(* 底辊采样反向 *)
	xMotRev_PrnRoller							: BOOL;(* 版辊电机反向运动 *)
	xSamRev_PrnRoller							: BOOL;(* 版辊采样反向 *)
	xMotRev_NetRoller							: BOOL;(* 网辊电机反向运动 *)

	xMotRev_NetRoller_Pressure_M				: BOOL;(* 网辊压力M侧电机反转/2021.11.16.133827/+4 *)
	xMotRev_NetRoller_Pressure_G				: BOOL;(* 网辊压力G侧电机反转 *)
	xMotRev_PrnRoller_Pressure_M				: BOOL;(* 版辊压力M侧电机反转 *)
	xMotRev_PrnRoller_Pressure_G				: BOOL;(* 版辊压力G侧电机反转 *)
	xMotRev_StrRoller_Pressure_M				: BOOL;(* 张带辊压力M侧电机反转 *)
	xMotRev_StrRoller_Pressure_G				: BOOL;(* 张带辊压力G侧电机反转 *)

	xFlag_RollerDn_BottomRoller					: BOOL;(* 底辊合压标志/底辊的胶辊 *)
	xFlag_RollerDn_PrnRoller					: BOOL;(* 印辊合压标志/靠上底辊 *)
	xFlag_RollerDn_NetRoller					: BOOL;(* 网辊合压标志/靠上版辊 *)

	xValid_BottomRoller							: BOOL;(* 底辊有效标志 *)
	iSid_BottomRoller							: INT;(* 底辊站id/初始-1/有效性通过查表确定 *)
	xStationOnline_BottomRoller					: BOOL;(* 站在线标志-底辊/读取站号以后实时更新 *)
	rAxisVel_BottomRoller						: REAL;(* 底辊轴速度 *)
(* 2021.12.29.152610/hdp *)

	xValid_PrnRoller							: BOOL;(* 印辊有效标志 *)
	iSid_PrnRoller								: INT;(* 版辊站id/初始-1/有效性通过查表确定 *)
	xStationOnline_PrnRoller					: BOOL;(* 站在线标志-版辊/读取站号以后实时更新 *)
	rAxisVel_PrnRoller							: REAL;(* 印版轴速度 *)

	xValid_NetRoller							: BOOL;(* 网辊有效标志 *)
	iSid_NetRoller								: INT;(* 网辊站id/初始-1/有效性通过查表确定 *)
	xStationOnline_NetRoller					: BOOL;(* 站在线标志-网辊/读取站号以后实时更新 *)
	rAxisVel_NetRoller							: REAL;(* 网辊轴速度 *)
(* 2021.12.29.152610/hdp *)

	iSid_PrnRoller_Pressure_M					: INT;(* 印辊压力电机M侧驱动器站号/初始-1 *)
	iSid_PrnRoller_Pressure_G					: INT;(* 印辊压力电机G侧驱动器站号/初始-1 *)
	iSid_PrnRoller_Pressure_2in1				: INT;(* 版辊压力电机驱动器站号 *)
		(*
		/2合1/初始-1
		/wCtlmod_PrnRoller_Pressure=2时用到 *)

	wCtlmod_NetRoller_Pressure					: WORD;(* 网辊压力控制方式 *)
		(*
		/0表示不控制(默认)
		/1为独立单轴控制
		/2为双轴控制
		/4为4轴驱动器控制 *)
	iSid_NetRoller_Pressure_M					: INT;(* 网辊压力电机M侧驱动器站号/初始-1 *)
	iSid_NetRoller_Pressure_G					: INT;(* 网辊压力电机G侧驱动器站号/初始-1 *)
	iSid_NetRoller_Pressure_2in1				: INT;(* 网辊压力电机驱动器站号 *)
		(*
		/2合1/初始-1
		/wCtlmod_NetRoller_Pressure=2时用到 *)

	iSid_Pressure_4in1							: INT;(* 压力电机4合1驱动器站号/版辊+网辊/初始-1 *)
		(*
		/wCtlmod_PrnRoller_Pressure=wCtlmod_NetRoller_Pressure=4时用到 *)
	iSid_StrRoller_Pressure_M					: INT;(* 印辊压力电机M侧驱动器站号/初始-1 *)
	iSid_StrRoller_Pressure_G					: INT;(* 印辊压力电机G侧驱动器站号/初始-1 *)
	iSid_StrRoller_Pressure_2in1				: INT;(* 版辊压力电机驱动器站号 *)
		(*
		/2合1/初始-1
		/wCtlmod_PrnRoller_Pressure=2时用到 *)

	iAxisIdx_PrnRoller_Pressure_M				: INT;(* 轴索引-版辊压力电机M侧 *)
	iAxisIdx_PrnRoller_Pressure_G				: INT;(* 轴索引-版辊压力电机G侧 *)
		(*
		/wCtlmod_PrnRoller_Pressure=2或4时用到*)

	iAxisIdx_NetRoller_Pressure_M				: INT;(* 轴索引-网辊压力电机M侧 *)
	iAxisIdx_NetRoller_Pressure_G				: INT;(* 轴索引-网辊压力电机G侧 *)
		(*
		/wCtlmod_NetRoller_Pressure=2或4时用到*)

	iAxisIdx_StrRoller_Pressure_M				: INT;(* 轴索引-网辊压力电机M侧 *)
	iAxisIdx_StrRoller_Pressure_G				: INT;(* 轴索引-网辊压力电机G侧 *)
		(*
		/wCtlmod_StrRoller_Pressure=2或4时用到*)

(* 2021.12.23.154424/hdp *)
	rPos_press_dn_PrnRoller_Pressure_M_Hmi		: REAL;(* 根据坐标系界面显示变量-hmi/合压位置/版辊压力电机M侧/单位:mm *)
	rPos_press_dn_PrnRoller_Pressure_G_Hmi		: REAL;(* 根据坐标系界面显示变量-hmi/合压位置/版辊压力电机G侧/单位:mm *)
	rPos_press_up_PrnRoller_Pressure_M_Hmi		: REAL;(* 根据坐标系界面显示变量-hmi/离压位置/版辊压力电机M侧/单位:mm *)
	rPos_press_up_PrnRoller_Pressure_G_Hmi		: REAL;(* 根据坐标系界面显示变量-hmi/离压位置/版辊压力电机G侧/单位:mm *)
	rPos_load_unload_PrnRoller_Pressure_M_Hmi	: REAL;(* 根据坐标系界面显示变量-hmi/装卸辊位置/版辊压力电机M侧/单位:mm *)
	rPos_load_unload_PrnRoller_Pressure_G_Hmi	: REAL;(* 根据坐标系界面显示变量-hmi/装卸辊位置/版辊压力电机G侧/单位:mm *)
(* end/hdp *)

(* 2021.12.22.185301/hdp *)
	rPos_press_dn_NetRoller_Pressure_M_Hmi		: REAL;(* 根据坐标系界面显示变量-hmi/合压位置/网辊压力电机M侧/单位:mm *)
	rPos_press_dn_NetRoller_Pressure_G_Hmi		: REAL;(* 根据坐标系界面显示变量-hmi/合压位置/网辊压力电机G侧/单位:mm *)
	rPos_press_up_NetRoller_Pressure_M_Hmi		: REAL;(* 根据坐标系界面显示变量-hmi/离压位置/网辊压力电机M侧/单位:mm *)
	rPos_press_up_NetRoller_Pressure_G_Hmi		: REAL;(* 根据坐标系界面显示变量-hmi/离压位置/网辊压力电机G侧/单位:mm *)
	rPos_load_unload_NetRoller_Pressure_M_Hmi	: REAL;(* 根据坐标系界面显示变量-hmi/装卸辊位置/网辊压力电机M侧/单位:mm *)
	rPos_load_unload_NetRoller_Pressure_G_Hmi	: REAL;(* 根据坐标系界面显示变量-hmi/装卸辊位置/网辊压力电机G侧/单位:mm *)
(* end/hdp *)

(* replaced@2021.12.22.185435/hdp
	lrAbsEnc_PrnRoller_Pressure_M				: LREAL;(* 版辊压力电机绝对值位置M侧/实时值 *)
	lrAbsEnc_PrnRoller_Pressure_G				: LREAL;(* 版辊压力电机绝对值位置G侧/实时值 *)
	lrAbsEnc_NetRoller_Pressure_M				: LREAL;(* 网辊压力电机绝对值位置M侧/实时值 *)
	lrAbsEnc_NetRoller_Pressure_G				: LREAL;(* 网辊压力电机绝对值位置G侧/实时值 *)
with... *)

(* 2021.12.22.185539/hdp *)
	rPos_PrnRoller_Pressure_M					: REAL;(* 版辊压力电机位置M侧/实时值|mm-根据坐标系变化 *)
	rPos_PrnRoller_Pressure_G					: REAL;(* 版辊压力电机位置G侧/实时值|mm-根据坐标系变化 *)
	rPos_NetRoller_Pressure_M					: REAL;(* 网辊压力电机位置M侧/实时值|mm-根据坐标系变化 *)
	rPos_NetRoller_Pressure_G					: REAL;(* 网辊压力电机位置G侧/实时值|mm-根据坐标系变化 *)
	rFrontSurfacePos_PrnRoller_Pressure_M		: REAL;(* 版辊压力电机M侧前表面位置|mm-根据坐标系变化 *)
	rFrontSurfacePos_PrnRoller_Pressure_G		: REAL;(* 版辊压力电机G侧前表面位置|mm-根据坐标系变化 *)
	rRearSurfacePos_PrnRoller_Pressure_M		: REAL;(* 版辊压力电机M侧后表面位置|mm-根据坐标系变化 *)
	rRearSurfacePos_PrnRoller_Pressure_G		: REAL;(* 版辊压力电机G侧后表面位置|mm-根据坐标系变化 *)
	rFrontSurfacePos_NetRoller_Pressure_M		: REAL;(* 网纹辊压力电机M侧前表面位置|mm-根据坐标系变化 *)
	rFrontSurfacePos_NetRoller_Pressure_G		: REAL;(* 网纹辊压力电机G侧前表面位置|mm-根据坐标系变化 *)
	rRearSurfacePos_NetRoller_Pressure_M		: REAL;(* 网纹辊压力电机M侧后表面位置|mm-根据坐标系变化 *)
	rRearSurfacePos_NetRoller_Pressure_G		: REAL;(* 网纹辊压力电机G侧后表面位置|mm-根据坐标系变化 *)
	xReConfirmPos0_AbsEnc						: BOOL;(*重新确认零位标志|由于机械位置或者电机位置跑了引起的异常需要重新确认零位 *)
	byTarPos_Roller									: BYTE;(*辊子目标位置|0 换版位
																		  1 离压位
																		  2 合压位*)
	byCurPos_Roller									: BYTE;(*辊子当前位置|0 换版位
																		  1 离压位
																		  2 合压位*)
	byInPos_Roller									: BYTE;(*辊子到位标志|.0 全部到位
																		  .1 版辊操作侧到位
																		  .2 版辊传动侧到位
																		  .3 网辊操作侧到位
																		  .4 网辊传动侧到位*)

	rPos_StrRoller_Pressure_M					: REAL;(* 张带辊压力电机位置M侧/实时值|mm-根据坐标系变化 *)
	rPos_StrRoller_Pressure_G					: REAL;(* 张带辊压力电机位置G侧/实时值|mm-根据坐标系变化 *)

(* 2021.12.23.154050/hdp *)

(* 2021.12.22.184937/hdp *)
	xMotEn_PrnRoller_Pressure					: BOOL;(* 版辊压力电机使能 *)
	xMotEn_NetRoller_Pressure					: BOOL;(* 网纹辊压力电机使能 *)
	xMotStop_PrnRoller_Pressure					: BOOL;(* 版辊压力电机停止 *)
	xMotStop_NetRoller_Pressure					: BOOL;(* 网纹辊压力电机停止 *)
	xNetRollSyncMoveByPrnRoll_Pressure			: BOOL;(* 网纹辊随版辊同时运动标志 *)
	rMoveDis_PrnRoller_Pressure_M				: REAL;(* 版辊压力操作侧运动距离|mm *)
	rMoveDis_PrnRoller_Pressure_G				: REAL;(* 版辊压力传动侧运动距离|mm *)
	rMoveDis_NetRoller_Pressure_M				: REAL;(* 网纹辊压力操作侧运动距离|mm *)
	rMoveDis_NetRoller_Pressure_G				: REAL;(* 网纹辊压力传动侧运动距离|mm *)
	xPosDevLarge_PrnRoller_Pressure				: BOOL;(* 版辊压力电机位置左右偏差太大 *)
	xPosDevLarge_NetRoller_Pressure				: BOOL;(* 网纹辊辊压力电机位置左右偏差太大 *)
	xTooClose_PrnRollerAndNetRoller_M			: BOOL;(* 版辊压力电机和网纹辊电机操作侧距离太近 *)
	xTooClose_PrnRollerAndNetRoller_G			: BOOL;(* 版辊压力电机和网纹辊电机传动侧距离太近 *)
	xSyncMoving_PrnRollAndNetRoll				: BOOL;(* 版辊和网辊同步运动中标志/2021.12.23.153947/lyt *)
	byCoordinate								: BYTE := 1;(* 坐标系类型选择:默认是使用网纹辊/0-使用各自坐标系/1-使用网纹辊坐标系|2-使用版辊坐标系 *)
	rCoordinateInter_PrnRollerAndNetRoller		: REAL;(* 版辊和网纹辊坐标系间隔|mm *)

(* end/hdp *)

	dwAxisAlrSts_NetRoller_Pressure_M			: DWORD;(* 网辊压力M侧报警状态 *)
	dwAlrCode_NetRoller_Pressure_M				: DWORD;(* 网辊压力M侧报警代码 *)
	dwAxisAlrSts_NetRoller_Pressure_G			: DWORD;(* 网辊压力G侧报警状态 *)
	dwAlrCode_NetRoller_Pressure_G				: DWORD;(* 网辊压力G侧报警代码 *)
	dwAxisAlrSts_PrnRoller_Pressure_M			: DWORD;(* 版辊压力M侧报警状态 *)
	dwAlrCode_PrnRoller_Pressure_M				: DWORD;(* 版辊压力M侧报警代码 *)
	dwAxisAlrSts_PrnRoller_Pressure_G			: DWORD;(* 版辊压力G侧报警状态 *)
	dwAlrCode_PrnRoller_Pressure_G				: DWORD;(* 版辊压力G侧报警代码 *)

(* 2021.12.23.153614/hdp *)
	byStsRapidAdjust							: BYTE;(* 快速对版状态|0不动作/1执行离开合压位动作/2合压位离开完成 *)
(* end/hdp *)

(*	//重新整理，按照每一个DWORD代表一种类型的辊子，目前有版辊网棍张带辊
	dwPressureMotor_Move						: DWORD;(* 色组压力电机控制按钮/可能来自实体/可能来自通讯及UI部分 *)
(*												/bit.0 : 印刷版辊M侧电机前进 *)
(*												/bit.1 : 印刷版辊M侧电机后退 *)
(*												/bit.2 : 印刷版辊G侧电机前进 *)
(*												/bit.3 : 印刷版辊G侧电机后退 *)
(*												/bit.4 : 印刷版辊压力电机前进 *)
(*												/bit.5 : 印刷版辊压力电机后退 *)
(*												/bit.6~7: 空闲 *)
(*												/bit.8 : 网辊M侧电机前进 *)
(*												/bit.9 : 网辊M侧电机后退 *)
(*												/bit.10: 网辊G侧电机前进 *)
(*												/bit.11: 网辊G侧电机后退 *)
(*												/bit.12: 网辊压力电机前进 *)
(*												/bit.13: 网辊压力电机后退 *)
(*												/bit.14~15: 空闲 *)
(*												/bit.16: 色组版辊压力电机前进 *)
(*												/bit.17: 色组版辊压力电机后退 *)
(*												/bit.18: 色组版辊压力电机合压 *)
(*												/bit.19: 色组版辊压力电机离压 *)
(*												/bit.20~23: 空闲 *)
(*												/bit.24: 色组版辊压力电机合压位确认按钮 *)
(*												/bit.25: 色组版辊压力电机离压位确认按钮 *)
(*												/bit.26: 色组版辊压力电机装版位确认按钮 *)
(*												/bit.27: 色组版辊压力电机零位确认按钮 *)
(*												/bit.28: 色组版辊压力电机边界位确认按钮 *)
(*												/bit.29~31: 空闲 *)

	dwPressureMotor_Move_II						: DWORD;(* 色组压力电机控制按钮/可能来自实体/可能来自通讯及UI部分 *)
(*												/bit.0 : 印刷张带辊M侧电机前进 *)
(*												/bit.1 : 印刷张带辊M侧电机后退 *)
(*												/bit.2 : 印刷张带辊G侧电机前进 *)
(*												/bit.3 : 印刷张带辊G侧电机后退 *)
(*												/bit.4 : 印刷张带辊压力电机前进 *)
(*												/bit.5 : 印刷张带辊压力电机后退 *)
(*												/bit.6~7: 空闲 *)
(*												/bit.8 : 色组网辊压力电机合压位确认按钮 *)
(*												/bit.9 : 色组网辊压力电机离压位确认按钮 *)
(*												/bit.10: 色组网辊压力电机装版位确认按钮 *)
(*												/bit.11: 色组网辊压力电机零位确认按钮 *)
(*												/bit.12: 色组网辊压力电机边界位确认按钮 *)
(*												/bit.13~15:空闲*)
(*												/bit.16: 色组张带辊压力电机合压位确认按钮 *)
(*												/bit.17: 色组张带辊压力电机离压位确认按钮 *)
(*												/bit.18: 色组张带辊压力电机装版位确认按钮 *)
(*												/bit.19: 色组张带辊压力电机零位确认按钮 *)
(*												/bit.20: 色组张带辊压力电机边界位确认按钮 *)
(*												/bit.21~23: 空闲 *)
(*												/bit.24: 色组网辊压力电机前进 *)
(*												/bit.25: 色组网辊压力电机后退 *)
(*												/bit.26: 色组网辊压力电机合压 *)
(*												/bit.27: 色组网辊压力电机离压 *)
(*												/bit.28: 色组张带辊压力电机前进 *)
(*												/bit.29: 色组张带辊压力电机后退 *)
(*												/bit.30: 色组张带辊压力电机合压 *)
(*												/bit.31: 色组张带辊压力电机离压 *)
*)

//重新整理，按照每一个DWORD代表一种类型的辊子，目前有1:版辊;	2:网棍;	3:张带辊
	adwPressureMotor_Move						: ARRAY[1..3] OF DWORD ;(* 色组压力电机控制按钮/可能来自实体/可能来自通讯及UI部分 *)
(*												/bit.0 : 辊M侧电机前进 *)
(*												/bit.1 : 辊M侧电机后退 *)
(*												/bit.2 : 辊G侧电机前进 *)
(*												/bit.3 : 辊G侧电机后退 *)
(*												/bit.4 : 辊压力电机前进 *)
(*												/bit.5 : 辊压力电机后退 *)
(*												/bit.6 : 辊压力电机长步持续前进 *)
(*												/bit.7 : 辊压力电机长步持续后退 *)
(*												/bit.8 : 辊压力电机离压 *)
(*												/bit.9 : 辊压力电机换版 *)
(*												/bit.10: 辊压力电机合压 *)
(*												/bit.11: 机械操作面板控制的印版辊压力电机换版走离压 *)
(*												/bit.12: 机械操作面板控制的印版辊压力电机离压走换版 *)
(*												/bit.13: 机械操作面板控制的印版辊压力电机在走离压换版的过程中停止 *)
//2026.02.23.132846
(*												/bit.14: 自动换版 *)
(*												/bit.15: 换版完成 *)
(*												/bit.16: 色组版辊压力电机合压位确认按钮 *)
(*												/bit.17: 色组版辊压力电机离压位确认按钮 *)
(*												/bit.18: 色组版辊压力电机装版位确认按钮 *)
(*												/bit.19: 显示换版状态 *)
(*												/bit.20~23: 空闲 *)
(*												/bit.24~31: 空闲 *)

	iCTL_Sample									: INT;(* 采样控制标志/ctl *)
	(*
	/以下时和套色有关的定义 *)
	iSampleCfgParam_ctl				:INT ;(*采样控制参数里的ctl		*)
	byColorIdCurrent				:BYTE;(*当前色序				*)
//	byColorIdFollow					:BYTE;(*跟踪色序				*)
	iRoundSampleDataSa							: INT;(* 粗采样数据起点 *)
	iRoundSampleViewDensity						: INT;(* 波形显示横向放大用的系数 *)
	byArcSts									: BYTE;(* 套色状态/bit0=报警/bit1=丢失 *)

(* 2021.12.6.145203/hdp/弃用.bit31的分配/单标记确认的操作通过主站和从站的界面提交动作/程序重新处理rOMKPos0_进行上下位机的同步即可 *)
(*												/bit31.单标记误差确认/状态改变1次认为操作1次/开机上电置位FALSE/2021.11.19.135306/+ *)

	wSts_TowardsTar_H							: WORD;(* 横向目标值状态 *)
	iPos_TowardsTar_H							: INT;(* 横向目标值运动位置实时值 *)
	dwSpecialRequest							: DWORD;(* 特殊请求位 *)
(*												/bit0.横向左-1 *)
(*												/bit1.横向左-2 *)
(*												/bit2.横向右-1 *)
(*												/bit3.横向右-2 *)
	dwExtendedMask								: DWORD;(* 扩展标志位 *)
(*												/bit0.色组记录粗采样数据/@2021.11.17.115203 *)
(*												/bit1.色组记录精采样数据/@2021.11.17.135352 *)
(*												/ *)
(*												/bit31.让料头/@2021.11.17.160031 *)

	rOMKPos0_									: REAL;(* 单标记0位 *)

	(* 色组调整相关 *)
	axCurCycleAdjustVal_Auto_done_vh			: ARRAY [1..2] OF BOOL;(* 本周期的自动套色调整消耗完成/[1]纵向/[2]横向 *)
	alrCurCycleAdjustVal_Auto_vh				: ARRAY [1..2] OF LREAL;(* 自动调整/[1]纵向/[2]横向 *)
	alrTotalAdjustVal_Auto_vh					: ARRAY [1..2] OF LREAL;(* 自动调整仓库/[1]纵向/[2]横向 *)
	alrExecutedAdjVal_Auto_vh					: ARRAY [1..2] OF LREAL;(* 已经执行的自动调整量/[1]纵向/[2]横向 *)

	axCurCycleAdjustVal_Rapid_done_vh			: ARRAY [1..2] OF BOOL;(* 本周期的快速对版调整消耗完成/[1]纵向/[2]横向 *)
	alrCurCycleAdjustVal_Rapid_vh				: ARRAY [1..2] OF LREAL;(* 快速对版调整/[1]纵向/[2]横向 *)
	alrTotalAdjustVal_Rapid_vh					: ARRAY [1..2] OF LREAL;(* 快速对版仓库/[1]纵向/[2]横向 *)
	alrExecutedAdjVal_Rapid_vh					: ARRAY [1..2] OF LREAL;(* 已经执行的快速调整量/[1]纵向/[2]横向 *)

	axCurCycleAdjustVal_ManuCoarse_done_vh		: ARRAY [1..2] OF BOOL;(* 本周期的手动粗调消耗完成/[1]纵向/[2]横向 *)
	alrCurCycleAdjustVal_ManuCoarse_vh			: ARRAY [1..2] OF LREAL;(* 手动粗调/[1]纵向/[2]横向 *)
	alrTotalAdjustVal_ManuCoarse_vh				: ARRAY [1..2] OF LREAL;(* 手动粗调仓库/[1]纵向/[2]横向 *)
	alrExecutedAdjVal_ManuCoarse_vh				: ARRAY [1..2] OF LREAL;(* 已经执行的手动粗调量/[1]纵向/[2]横向 *)

	axCurCycleAdjustVal_ManuFine_done_vh		: ARRAY [1..2] OF BOOL;(* 本周期的手动细调消耗完成/[1]纵向/[2]横向 *)
	alrCurCycleAdjustVal_ManuFine_vh			: ARRAY [1..2] OF LREAL;(* 手动细调/[1]纵向/[2]横向 *)
	alrTotalAdjustVal_ManuFine_vh				: ARRAY [1..2] OF LREAL;(* 手动细调仓库/[1]纵向/[2]横向 *)
	alrExecutedAdjVal_ManuFine_vh				: ARRAY [1..2] OF LREAL;(* 已经执行的手动细调量/[1]纵向/[2]横向 *)

	axCurCycleAdjustVal_Coupling_done_vh		: ARRAY [1..2] OF BOOL;(* 本周期的耦合消耗完成/[1]纵向/[2]横向 *)
	alrCurCycleAdjustVal_Coupling_vh			: ARRAY [1..2] OF LREAL;(* 耦合量/[1]纵向/[2]横向 *)
	alrTotalAdjustVal_Coupling_vh				: ARRAY [1..2] OF LREAL;(* 耦合量仓库/[1]纵向/[2]横向 *)
	alrExecutedAdjVal_Coupling_vh				: ARRAY [1..2] OF LREAL;(* 已经执行的耦合量/[1]纵向/[2]横向 *)

(* 2021.12.30.165518/lyt/+ *)
	tMovingTimeSa									:TIME;(*运动启动时间|ms*)
	xAutoSts_Roller_Pressure						:BOOL;(*压力辊自动状态*)

	(*
	/保留部分 *)
	xMoveEnable_Motor						: BOOL;(*电机运动使能|用于控制驱动器是否进行电机控制|与单联动比较切换电机是否运动*)
	byHandWheelSts: BYTE;(**)

	rCurrent_PrnPressure_M: REAL;//版辊M侧电机电流
	rCurrent_PrnPressure_G: REAL;//版辊M侧电机电流
	rCurrent_NetPressure_M: REAL;//网辊M侧电机电流
	rCurrent_NetPressure_G: REAL;//网辊M侧电机电流
	rCurrent_StrPressure_M: REAL;//张带辊M侧电机电流
	rCurrent_StrPressure_G: REAL;//张带辊M侧电机电流
	wSts_HorzManuPreReg						: WORD; (* 横向手动预套准状态标志|bit0运行标志|bit1正转|bit2反转|bit3左限位|bit4右限位|bit5停止 *)
	iPos_HorzManuPreReg						: INT;(*横向手动预套准位置|*)
	xFlag_HorzPreRegister_ing				: BOOL;(*横向预套准进行中|*)
	xFlag_HorzPreRegister_end				: BOOL;(*横向预套准完成|*)

	diPreReg_RepeatVal_H					: DINT;(*预套准重复值-横向|单位:mm|*)
	diPreReg_SetupVal_H						: DINT;(*预套准设定值-横向|单位:mm|*)

	lrVelocity_CoatingPrn					: LREAL;(*涂布速度|*)
	byBtn_AdjModeSwitch_CoatingPrn			: BYTE;(*涂布调整方式切换按钮|*)
	xAxisInching							: BOOL;(*版辊单运行中*)
	xAxisInching_Net						: BOOL;(*网辊单运行中*)
	iPhase_InstallPlate						: INT;(*装版相位|*)
	iPhase_RegisterOk						: INT;(*套准相位|版套印准确的相位<通用相位和相位保存/恢复都可以复用该变量>|*)
	//lrPreReg_ConstVal						: LREAL;(*预套准色组间固定料长部分|单位:mm*)

	xEn_Motor_PrnRoller						: BOOL;(*版辊开始运行标志-运动过程中序保证该标志一直有效*)
	xEn_Motor_NetRoller						: BOOL;(*网辊开始运行标志-运动过程中序保证该标志一直有效*)
	xEn_Motor_BottomRoller						: BOOL;(*底辊开始运行标志-运动过程中序保证该标志一直有效*)

	xFlag_FastAdjusting						: BOOL;//快速对半中2023.8.18.104925新增标志
	xFlag_MediumAdjusting				: BOOL;//粗调中
	xFlag_SlowAdjusting				: BOOL;//细调/等

	//以下位色组各轴的离线报警位置偏差报警标志
	xNetOffline_Horz:BOOL;
	xAxisAlarm_Horz:BOOL;
	xPosDeviationAlarm_Horz:BOOL;

	xNetOffline_PrnRoller:BOOL;
	xAxisAlarm_PrnRoller:BOOL;
	xPosDeviationAlarm_PrnRoller:BOOL;

	xNetOffline_NetRoller:BOOL;
	xAxisAlarm_NetRoller:BOOL;
	xPosDeviationAlarm_NetRoller:BOOL;

	xNetOffline_BottomRoller:BOOL;
	xAxisAlarm_BottomRoller:BOOL;
	xPosDeviationAlarm_BottomRoller:BOOL;

	xNetOffline_Prn_Pressure_M:BOOL;
	xAxisAlarm_Prn_Pressure_M:BOOL;
	xPosDeviationAlarm_Prn_Pressure_M:BOOL;

	xNetOffline_Prn_Pressure_G:BOOL;
	xAxisAlarm_Prn_Pressure_G:BOOL;
	xPosDeviationAlarm_Prn_Pressure_G:BOOL;

	xNetOffline_Net_Pressure_M:BOOL;
	xAxisAlarm_Net_Pressure_M:BOOL;
	xPosDeviationAlarm_Net_Pressure_M:BOOL;

	xNetOffline_Net_Pressure_G:BOOL;
	xAxisAlarm_Net_Pressure_G:BOOL;
	xPosDeviationAlarm_Net_Pressure_G:BOOL;

	xNetOffline_Str_Pressure_M:BOOL;
	xAxisAlarm_Str_Pressure_M:BOOL;
	xPosDeviationAlarm_Str_Pressure_M:BOOL;

	xNetOffline_Str_Pressure_G:BOOL;
	xAxisAlarm_Str_Pressure_G:BOOL;
	xPosDeviationAlarm_Str_Pressure_G:BOOL;

	xNetOffline_PHOTOCELL:BOOL;
	xAxisAlarm_PHOTOCELL:BOOL;
	xPosDeviationAlarm_PHOTOCELL:BOOL;
	//2023.8.18.143436各个轴的具体报警信息；

	dwAlarmDetail_Prn:DWORD;//轴报警信息-版辊
	dwAlarmDetail_Net:DWORD;//轴报警信息-wnag辊
	dwAlarmDetail_Bottom:DWORD;//轴报警信息-底辊
	dwAlarmDetail_Prn_M:DWORD;//轴报警信息-版辊_M
	dwAlarmDetail_Prn_G:DWORD;//轴报警信息-版辊_G
	dwAlarmDetail_Net_M:DWORD;//轴报警信息-网辊_M
	dwAlarmDetail_Net_G:DWORD;//轴报警信息-网辊_G
	dwAlarmDetail_Horz:DWORD;//轴报警信息-横向
	dwAlarmDetail_PHOTOCELL:DWORD;//光电眼
	dwAlarmDetail_Str_M:DWORD;//轴报警信息-网辊_M
	dwAlarmDetail_Str_G:DWORD;//轴报警信息-网辊_G

	xOnline_NR_M_: BOOL;(* 网辊压力M侧在线 *)
	xOnline_NR_G_: BOOL;(* 网辊压力G侧在线 *)
	xOnline_PR_M_: BOOL;(* 版辊压力M侧在线 *)
	xOnline_PR_G_: BOOL;(* 版辊压力G侧在线 *)
	xOnline_STR_M_: BOOL;(* 版辊压力M侧在线 *)
	xOnline_STR_G_: BOOL;(* 版辊压力G侧在线 *)

	iSid_Horiz_: INT;(* 横向伺服站点 *)
	xMotRev_Horiz_: BOOL;(* 横向伺服反转 *)
	xOnline_Horiz_: BOOL;(* 横向伺服在线 *)
	rErr_V:REAL;
	rErr_H:REAL;

	xValid_PhotoCell							: BOOL;		(* 光电眼有效标志 *)
	iSid_PhotoCell							: INT;			(* 光电眼站id/初始-1/有效性通过查表确定 *)
	xStationOnline_PhotoCell					: BOOL;		(* 站在线标志-光电眼/读取站号以后实时更新 *)
	xMotRev_PhotoCell							: BOOL;		(* 光电眼电机反向运动 *)
	rAxisVel_PhotoCell						: REAL;			(* 光电眼轴速度 *)

(*2023.9.25.135838*)
	byEn_Motor_Pressure_: BYTE;
	//每个色组可以有8个龙门控制轴-4组，目前只用到了4个
	byEn_Motor_Trap_: BYTE;(*.0 横向
							 .1	光电眼*)
	//每个色组可以有8个点位控制轴-4组，目前只用到了1个，横向，其他当预留吧，反正一个BOOL和一个BYTE是一样的；
(*2023.10.27.085455*)
	//横向软限位
(*
	lrLimit_Left : LREAL;
	lrLimit_Right : LREAL;
*)
	abyRsv_Data1: ARRAY [1..16] OF BYTE;
	rweigth_Prn_Bottom_Cur					: REAL;//这个是版辊中心到版辊和底辊/中心辊切点的横向距离
	rweigth_Prn_Net_Cur					: REAL;//这个是版辊中心到版辊和网辊切点的横向距离
	rweigth_Net_Prn_Cur				: REAL;//这个是网辊中心到网辊与版辊切点的横向距离
	rweigth_Net_Load_Cur					: REAL;//这个是版辊中心到版辊和网辊切点的横向距离

	//bai.zy | 2024.04.03.132443 | 光电眼软限位位置记录
	lrPhotoCellPosLimit_M : LREAL;
	lrPhotoCellPosLimit_G : LREAL;

(*2023.10.14.105907加热部分增加|28zijie*)
(*加热相关*)
(* 加热部分 *)
	rPV_UnitTemCtl							: REAL;(* 色组温度控制实时值 *)

(* 刮刀部分 *)

	rHz_UnitExhaust_CurrRD					: REAL;(* 排风当前回读频率/pdu上行给主站/ *)
	rHz_UnitExhaust_CurrWR					: REAL;(* 排风当前写入频率/pdu下行给从站/ *)
	wSTS_UnitExhaust						: WORD;(* 排风状态|/.0 通讯返回运行状态
												   /.6 排风打开超时-
												   /.7 485通讯断开标志
												   高8位作为报警码*)
	dwCtlBits_UnitBaseCraft					: DWORD;(* 用户基础工艺控制位/加热/递墨辊/刮刀/热风 *)
												(*
												/ .bit0 ~bit3  刮刀
												/	/.bit0 刮刀自动(TRUE)/手动(FALSE)
												/	/.bit1 刮刀开(TRUE)/关(FALSE)
												/	/.bit2 刮刀运行信号/控制变频器启动
												/	/.bit3
												/ .bit4 ~bit7  递墨辊
												/	/.bit4 递墨辊自动(TRUE)/手动(FALSE)
												/	/.bit5 递墨辊正转(TRUE)/关或反转(FALSE)
												/	/.bit6 递墨辊反转(TRUE)/关或正转(FALSE)
												/	/.bit7 递墨辊运行信号/控制变频器启动-与/.4/.5共同确定正转还是反转
												/ .bit8 ~bit11 热风I
												/	/.bit8 热风I开(TRUE)/关(FALSE)
												/	/.bit9 热风I运行信号/控制变频器启动
												/	/.bit10
												/	/.bit11
												/ .bit12~bit15 热风II
												/	/.bit12 热风II开(TRUE)/关(FALSE)
												/	/.bit13 热风II运行信号/控制变频器启动
												/	/.bit14
												/	/.bit15
												/ .bit16~bit23
												/	/ .bit16 加热方式（水）
												/	/ .bit17 加热方式（电）
												/	/ .bit18 I档
												/	/ .bit19 II档
												/	/ .bit20 III档
												/	/ .bit21
												/	/ .bit22
												/ .bit23~bit26
												/	/ .bit23 刮刀故障复位
												/	/ .bit24 递墨故障复位
												/	/ .bit25 热风I故障复位
												/	/ .bit26 热风II故障复位
												/   / .bit27 排风故障复位
												/ .bit28~bit31 /2022.3.23.152646/hdp/预分配好/为和界面作绑定
												/	/ .bit28 排风开(TRUE)/关(FALSE)
												/	/ .bit29 排风运行信号/控制变频器启动
												/	/ .bit30
												(*2022.4.20.091641 移动到此处*)
												/	/ .bit31: 2022.4.20.091632|冷风机开关使能位||
												*)
	lrAxisScraperVel						: LREAL;(*刮刀速度输出|*)
	rAI0Value_16D							: REAL;(*16D io接口获取的模拟量输入值|*)
	rTempValue_16D							: REAL;(*16D io接口获取的温度值|*)
	rAO0Value_16D							: REAL;(*16D io接口输出的电压值1|*)
	rAO1Value_16D							: REAL;(*16D io接口输出的电压值2|*)
	rDemarcate_Read_1					: REAL;
	rDemarcate_Read_2					: REAL;
	rDemarcate_Write_1					: REAL;
	rDemarcate_Write_2					: REAL;

	//2023.11.21.155350色组压印到压印的料长
	lrArc_length_PrintPoint				: LREAL;
	dwSlaveBtn_HMI:DWORD;
												(*2023.12.22.205559
												bit0:纵向上调；
												bit1:纵向下调；
												bit2:横向左调；
												bit3:横向右调；
												bit4:版辊M侧前进；
												bit5:版辊M侧后退；
												bit6:版辊平行前进；
												bit7:版辊平行后退；
												bit8:版辊G侧前进；
												bit9:版辊G侧后退；
												bit10:网辊M侧前进；
												bit11:网辊M侧后退；
												bit12:网辊平行前进；
												bit13:网辊平行后退；
												bit14:网辊G侧前进；
												bit15:网辊G侧后退；

												*)
//秦华带长调整开关
	xAdjBandLen							 : BOOL;

	// 2024.10.21.114937 | bai.zy | 版辊网辊操作侧传动侧标定平行标志、标定平行后产生的误差值 15字节
	xConfirmParallelPos_Prn : BOOL;//平行确认按钮
	xConfirmParallelPos_Net : BOOL;
	xConfirmParallelPos_Str : BOOL;
	rParallelError_Prn_MM : REAL;//计算出的两侧误差
	rParallelError_Net_MM : REAL;
	rParallelError_Str_MM : REAL;

//根据单圈绝对值计算的装版位置；2024.10.22.222722	4字节
	diPhase_Enc_InstallPlate: DINT;

//2024.12.03.162342 | 增加调试阶段的压力运动 ，标定最大限位  ---3字节
	axCalidPressLimit_Max : ARRAY[1..3] OF BOOL;

	wUnit_input_I : WORD;
						(*
							bit0: 联动
							bit1: 单运行
							bit2: 急停输入
							bit3: 报警
							bit4: 细调
							bit5: 自动合压
							bit6: 合压输入
							bit7: 离压输入
							bit8: 点动离压
							bit9: 纵向上
							bit10: 纵向下
							bit11: 横向左限位
							bit12: 横向左
							bit13:
							bit14:
							bit15: IO监控标志位
						*)
	wUnit_input_II : WORD;
							(*
							bit0: 横向右
							bit1: 横向右限位
							bit2: 横向电机快
							bit3: 冷风开关
							bit4: 冷风按钮
							bit5: 热风报警
							bit6: 热风开关
							bit7: 热风按钮
							bit8: 温度到达预设
							bit9: 加热I档
							bit10:加热II档
							bit11:加热III档
							bit12: 加热按钮
						*)
	wUnit_input_III : WORD;
						(*
							bit0: 刮刀变频报警
							bit1: 刮刀开关
							bit2: 排风开关
							bit3: 递墨辊正转
							bit4: 递墨辊上
							bit5: 排风按钮
							bit6: 加速
							bit7: 减速
							bit8: 停机
							bit9: 快停
							bit10: PTC过温
							bit11: 顶板送
						*)
	wUnit_output_I : WORD;
						(*
							bit0: 联动指示
							bit1: 单运行指示
							bit2: 急停灯输出
							bit3: 套色正常
							bit4: 套色报警
							bit5: 套色丢失
							bit6: 横向正转输出
							bit7: 本组套色报警
							bit8: 合压输出
							bit9: 横向反转输出
							bit10: 轴故障指示
							bit11: 离压输出
							bit12: 冷风输出
						*)
	wUnit_output_II : WORD;
						(*
							bit0: 热风输出
							bit1: 色组排风输出
							bit2: 加热I输出
							bit3: 加热II输出
							bit4: 加热III输出
							bit5: 刮刀使能
							bit6: 递墨辊正转
							bit7: 递墨辊上
						*)
	rHz_UnitHotWind2_CurrRD					: REAL;(* 热风当前回读频率/pdu上行给主站/ *)
	rHz_UnitHotWind2_CurrWR					: REAL;(* 热风当前写入频率/pdu下行给从站/ *)
	wSTS_UnitHotWind_2						: WORD;(* 热风II状态 *)
	rHz_UnitHotWind_CurrRD					: REAL;(* 热风当前回读频率/pdu上行给主站/ *)
	rHz_UnitHotWind_CurrWR					: REAL;(* 热风当前写入频率/pdu下行给从站/ *)
	wSTS_UnitHotWind						: WORD;(* 热风状态 |.0 运行\停止
												               /.6 热风风打开超时-
												  			   /.7 485通讯断开标志*)
	rHz_UnitScraper_CurrRD					: REAL;(* 刮刀当前回读频率/pdu上行给主站/ *)
	rHz_UnitScraper_CurrWR					: REAL;(* 刮刀当前写入频率/pdu下行给从站/ *)
	wSTS_UnitScraper						: WORD;(* 刮刀状态/pdu上行给主站/ |.0 运行\停止
												              				  /.6 刮刀打开超时-
												                              /.7 485通讯断开标志*)
	rHz_UnitInkRoller_CurrRD				: REAL;(* 递墨辊当前回读频率/pdu上行给主站/ *)
	rHz_UnitInkRoller_CurrWR				: REAL;(* 递墨辊当前写入频率/pdu下行给从站/ *)
	wSTS_UnitInkRoller						: WORD;(* 递墨辊状态/pdu上行给主站 |.0 运行\停止
												              				   /.6 递墨辊刀打开超时
												                               /.7 485通讯断开标志*)
	wSTS_UnitTemCtl							: WORD;(* 色组温度控制报警代码|低8位作为运行状态
																				/.0 通讯返回运行状态
																				/.1 加热使能输出状态
												  高8位作为报警状态/.8 断偶标志
																   /.9 超温标志
																   /.10 离线标志*)
	rVerror_Lp		: REAL;(*低通滤波以后的误差@误差平均值需要写0*)
	xArcErrValid		: BOOL;
	xArcErrValid_Use_Niu: BOOL;
	iArcErr_V: INT;(*套色的纵向误差@每圈更新一次并按bit置位表示误差有效*)
	xSkipHeader								: BOOL;(*让料头*)
	xSkipHeaderSts							: BOOL;(*让料头状态@每次接料都会计算@根据是否打开让料头标志是否输出xSkipHeader*)
	xArcErrIsValid_V						: BOOL;(*纵向误差有效*)
	xArcErrIsValid_H						: BOOL;(*横向误差有效*)
	(*套色相关一些值写入到轴参数中-50BYTES@2024.6.15.103803*)
	xArcErrIsLost_V							: BOOL;	(*纵向套色误差丢失*)
	xArcErrIsFake_V							: BOOL;	(*纵向套色误差飞点*)
	(*套色相关一些值写入到轴参数中-50BYTES@2024.6.15.103803*)
	xArcErrIsLost_H							: BOOL;	(*横向套色误差丢失*)
	xArcErrIsFake_H							: BOOL;	(*横向套色误差飞点*)

	xArcErrIsAlarm_V						: BOOL;(*纵向报警*)
	xArcErrIsAlarm_H						: BOOL;(*横向报警*)
	xFlag_PressDn							: BOOL;(*色组压辊标志*)
	iFinalAdjust_V							: INT;
	iFinalAdjust_H							: INT;

	iVerror_Follow1UnitByErrTrans			: INT;(*纵向误差跟踪第一色@通过传递计算值*)

	(*增加一下误差队列*)
	byIndex: BYTE;
	aiError_V_History: ARRAY [1..50] OF INT;(*纵向误差队列*)
	aiError_H_History: ARRAY [1..50] OF INT;(*横向误差队列*)

	(*新增参数|wang.nt|2025.08.08.155511*)
	alrCurcycleAdjustVal_Compensate_vh: ARRAY [1..2] OF LREAL; (* 补偿量*)
	alrTotalAdjustVal_Compensate_vh: ARRAY [1..2] OF LREAL; (* 补偿量仓库*)
	alrExecutedAdjVal_Compensate_vh: ARRAY [1..2] OF LREAL; (* 已经执行的补偿量*)
	axCurCycleAdjustVal_Compensate_done_vh: ARRAY [1..2] OF BOOL;
	xAxisAutoPressed					: BOOL;
	byRapidAdjustStep					: BYTE;
	xRapidAdjust_ing					: BOOL;
	iRapidAdjust_TimingCnt				: INT;
	(*新增工艺参数|2025.08.15.151756*)
	byFreq_ExhaustAir : BYTE;
	byFreqCur_ExhaustAir :BYTE ;
	byAirInletWindDoorValue_FeedBack : BYTE;

(*2025.8.19.201439新增||需要在main里面赋值一下*)
	uiFSampleCounter: UINT;
	iManualPlateAdjustment_disp: INT;(*2025.5.15.195937/han.dp/+单位mm@显示当前值*)
	iAdjValue_V								: INT;(*统计纵向总调整量-用于实现新型耦合方式@um*)
(*2025.8.22.212351*)
	lrEnc_Pos: LREAL;(*版辊编码器位置*)
(*2025.9.24.175237||从这里开始属于润新测试后新增变量，与家里参数不再一致，回去更新吧*)
	xAxisInf_IO_Alarm_HotBlower: BIT;(*风机变频故障*)
	xAxisInf_IO_Alarm_PowerAdj: BIT;(*功率调整器故障*)
	xAxisInf_IO_Alarm_HeatClose: BIT;(*加热电源脱开故障*)
	xAxisInf_IO_Alarm_HeatLimit: BIT;(*超温报警*)
	xAxisInf_IO_Alarm_InkRoller: BIT;(*递墨变频故障*)
	xAxisInf_IO_Alarm_Scraper: BIT;(*刮刀变频故障*)
	xAxisInf_IO_Alarm_ExhAir: BIT;(*排风变频故障*)
	xInValidVirtualCnt: BIT;(**)
	wVirTual_Cnt: WORD;(*虚拟码盘计数*)
	wVirTual_Sts: WORD;(*虚拟码盘状态*)
	lrPrf_Pos: LREAL;(*版辊编码器位置*)
	byEnableModeSwitchDne: BYTE;
	rAxisPrfVel: REAL;
	iAxisPrnRunCaseId: INT;

	//2026.5.9.190555+
	dwLockTime_GetArcErr:DWORD;(*获取到套色误差的锁存时间@华南理工需要*)
	dwTime_Lock:DWORD;//锁存时间
	dwEnc_Lock:DWORD;//锁存编码器
	iStationId_CTL:INT:=-1;//控制的站id@例如月光宝盒\月光宝盒站id,如果是16d则和iStationId保持一样(iStationId该变量现在是电机驱动器的站号注意)

	//xNetOffline_Ctl色组控制器离线
	xNetOffline_Ctl: BOOL;

END_STRUCT
END_TYPE

{IMPLEMENTATION}
